Fanuc KAREL source: KT00841.KL

PROGRAM KT00841
%NOLOCKGROUP
VAR
  B1: BOOLEAN
  B2: BOOLEAN
  OUT: REAL
BEGIN
  B1 = TRUE
  B2 = FALSE
  B1 = TRUE
  B2 = FALSE
  OUT = SQRT(B1)
END KT00841
